(* PLC project Mixer.project, CODESYS CODESYS V3.5 SP19 *)
(* stored: creationDateTime 2025-05-14T10:21:07.1872635, modificationDateTime 2025-05-14T10:20:51.4312196 *)

PROGRAM PLC_PRG
  VAR
    Start_PB AT %IX0.0 : BOOL;  (* Start pushbutton *)
    Stop_PB AT %IX0.1 : BOOL;  (* Stop pushbutton *)
    Motor_Fault AT %IX0.2 : BOOL;  (* Agitator motor overload *)
    Manual_Run AT %IX0.3 : BOOL;  (* Manual jog selector *)
    Agitator_Run AT %QX0.0 : BOOL;  (* Agitator contactor *)
    Batch_Done AT %QX0.1 : BOOL;  (* Batch complete lamp *)
  END_VAR
  VAR
    Bypass_Mode : BOOL;  (* Maintenance bypass *)
    Run_Request : BOOL;
    Mix_Timer : TON;
  END_VAR

            (* Mixer sequence *)
IF Start_PB AND NOT Bypass_Mode THEN
    Run_Request := TRUE;
END_IF
IF NOT Stop_PB OR Motor_Fault THEN
    Run_Request := FALSE;
END_IF

Mix_Timer(IN := Run_Request, PT := T#45S);
Agitator_Run := Run_Request AND NOT Mix_Timer.Q;

IF Bypass_Mode THEN
    Agitator_Run := Manual_Run;
END_IF

Batch_Done := Mix_Timer.Q;
          
END_PROGRAM

CONFIGURATION Device
  RESOURCE Application ON PLC
    TASK MainTask(INTERVAL := T#20ms, PRIORITY := 1);
    PROGRAM PLC_PRG WITH MainTask : PLC_PRG;
  END_RESOURCE
END_CONFIGURATION
